FUNCTION_BLOCK SEC_SWITCH_LR_QUARTER_LWORD (* Section-Switcher: Teilbreiten von links und von rechts abschalten, bis 32 Sections, Maske als LWORD im Condensed Work State (2 Bit je Section) *)
  (* Standard: 61499-2; Description: Copyright (c) 2026 Meisterschulen am Ostbahnhof This program and the accompanying materials are made available under the terms of the Eclipse Public License 2.0 which is available at https://www.eclipse.org/legal/epl-2.0/ SPDX-License-Identifier: EPL-2.0 *)
  (* Version 1.1, 2026-11-01, Franz Höpfinger, Meisterschulen am Ostbahnhof, Alle aus und eigener Zaehler 0: LEFT/RIGHT_OFF_DEC uebernimmt zuerst alle abgeschalteten Sections (nach ALL_OFF schaltet Links_Ein von rechts, Rechts_Ein von links zu) *)
  (* Version 1.0, 2026-10-31, Franz Höpfinger, Meisterschulen am Ostbahnhof, initial implementation *)
  PACKAGE logiBUS::sections;
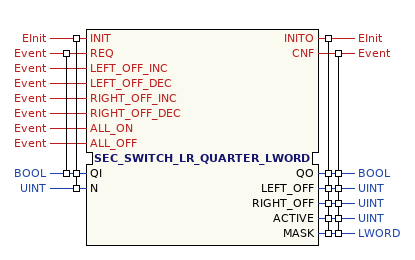
  EVENT_INPUT
    INIT : EInit WITH QI, N; (* Initialisierung, Zaehler auf 0 *)
    REQ WITH QI; (* Maske und Zaehler erneut ausgeben *)
    LEFT_OFF_INC; (* Von links eine Section mehr abschalten *)
    LEFT_OFF_DEC; (* Von links eine Section wieder zuschalten *)
    RIGHT_OFF_INC; (* Von rechts eine Section mehr abschalten *)
    RIGHT_OFF_DEC; (* Von rechts eine Section wieder zuschalten *)
    ALL_ON; (* Alle Sections zuschalten (beide Zaehler 0) *)
    ALL_OFF; (* Alle Sections abschalten (LEFT_OFF = N, RIGHT_OFF = 0) *)
  END_EVENT
  EVENT_OUTPUT
    INITO : EInit WITH QO, LEFT_OFF, RIGHT_OFF, ACTIVE, MASK; (* Initialisierung bestaetigt *)
    CNF WITH QO, LEFT_OFF, RIGHT_OFF, ACTIVE, MASK; (* Zaehler oder Maske neu berechnet *)
  END_EVENT
  VAR_INPUT
    QI : BOOL := TRUE; (* Nur an INIT und REQ: INIT+ aktiv, INIT- deaktiviert (Maske alle frei), REQ- ohne Wirkung *)
    N : UINT; (* Anzahl Sections (1..32, groesser wird auf 32 begrenzt) *)
  END_VAR
  VAR_OUTPUT
    QO : BOOL; (* TRUE = aktiv und Ereignis ausgefuehrt *)
    LEFT_OFF : UINT; (* Anzahl von links abgeschalteter Sections *)
    RIGHT_OFF : UINT; (* Anzahl von rechts abgeschalteter Sections *)
    ACTIVE : UINT; (* Anzahl freier Sections *)
    MASK : LWORD; (* Maske, 2 Bit je Section: 01 frei, 00 gesperrt, 11 nicht vorhanden (Section > N); Bits 1..0 = Section 1 (links) *)
  END_VAR
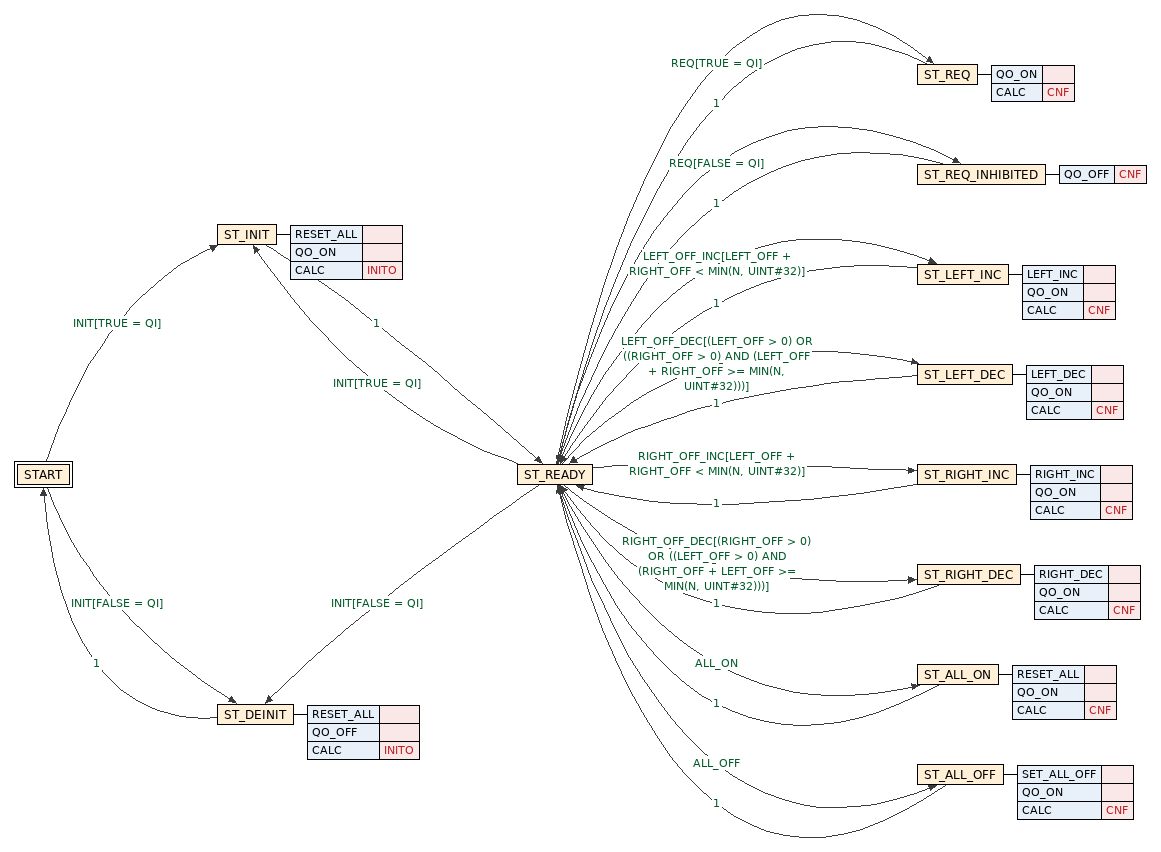
  EC_STATES
    START; (* Nicht initialisiert bzw. deaktiviert *)
    ST_INIT : RESET_ALL, QO_ON, CALC -> INITO; (* INIT+: N uebernehmen, Zaehler 0 *)
    ST_READY; (* Aktiv *)
    ST_DEINIT : RESET_ALL, QO_OFF, CALC -> INITO; (* INIT-: deaktiviert, Maske alle frei *)
    ST_REQ : QO_ON, CALC -> CNF; (* REQ+: Maske und Zaehler ausgeben *)
    ST_REQ_INHIBITED : QO_OFF -> CNF; (* REQ-: nichts aendern, nur melden *)
    ST_LEFT_INC : LEFT_INC, QO_ON, CALC -> CNF;
    ST_LEFT_DEC : LEFT_DEC, QO_ON, CALC -> CNF;
    ST_RIGHT_INC : RIGHT_INC, QO_ON, CALC -> CNF;
    ST_RIGHT_DEC : RIGHT_DEC, QO_ON, CALC -> CNF;
    ST_ALL_ON : RESET_ALL, QO_ON, CALC -> CNF;
    ST_ALL_OFF : SET_ALL_OFF, QO_ON, CALC -> CNF;
  END_STATES
  EC_TRANSITIONS
    START TO ST_INIT := INIT[TRUE = QI];
    START TO ST_DEINIT := INIT[FALSE = QI];
    ST_INIT TO ST_READY := 1;
    ST_DEINIT TO START := 1;
    ST_READY TO ST_INIT := INIT[TRUE = QI];
    ST_READY TO ST_DEINIT := INIT[FALSE = QI];
    ST_READY TO ST_REQ := REQ[TRUE = QI];
    ST_REQ TO ST_READY := 1;
    ST_READY TO ST_REQ_INHIBITED := REQ[FALSE = QI];
    ST_REQ_INHIBITED TO ST_READY := 1;
    ST_READY TO ST_LEFT_INC := LEFT_OFF_INC[LEFT_OFF + RIGHT_OFF < MIN(N, UINT#32)];
    ST_LEFT_INC TO ST_READY := 1;
    ST_READY TO ST_LEFT_DEC := LEFT_OFF_DEC[(LEFT_OFF > 0) OR ((RIGHT_OFF > 0) AND (LEFT_OFF + RIGHT_OFF >= MIN(N, UINT#32)))];
    ST_LEFT_DEC TO ST_READY := 1;
    ST_READY TO ST_RIGHT_INC := RIGHT_OFF_INC[LEFT_OFF + RIGHT_OFF < MIN(N, UINT#32)];
    ST_RIGHT_INC TO ST_READY := 1;
    ST_READY TO ST_RIGHT_DEC := RIGHT_OFF_DEC[(RIGHT_OFF > 0) OR ((LEFT_OFF > 0) AND (RIGHT_OFF + LEFT_OFF >= MIN(N, UINT#32)))];
    ST_RIGHT_DEC TO ST_READY := 1;
    ST_READY TO ST_ALL_ON := ALL_ON;
    ST_ALL_ON TO ST_READY := 1;
    ST_READY TO ST_ALL_OFF := ALL_OFF;
    ST_ALL_OFF TO ST_READY := 1;
  END_TRANSITIONS
  ALGORITHM RESET_ALL IN ST:
LEFT_OFF := 0;
RIGHT_OFF := 0;
  END_ALGORITHM
  ALGORITHM LEFT_INC IN ST:
LEFT_OFF := LEFT_OFF + 1;
  END_ALGORITHM
  ALGORITHM LEFT_DEC IN ST:
(* Alle aus und eigener Zaehler 0: diese Seite uebernimmt zuerst alle
   abgeschalteten Sections, damit beide Seiten nach ALL_OFF zuschalten *)
IF (LEFT_OFF = 0) AND (RIGHT_OFF > 0) AND (LEFT_OFF + RIGHT_OFF >= MIN(N, UINT#32)) THEN
	LEFT_OFF := RIGHT_OFF;
	RIGHT_OFF := 0;
END_IF;
(* Schutz gegen UINT-Unterlauf, zusaetzlich zur ECC-Bedingung *)
IF LEFT_OFF > 0 THEN
	LEFT_OFF := LEFT_OFF - 1;
END_IF;
  END_ALGORITHM
  ALGORITHM RIGHT_INC IN ST:
RIGHT_OFF := RIGHT_OFF + 1;
  END_ALGORITHM
  ALGORITHM RIGHT_DEC IN ST:
(* Alle aus und eigener Zaehler 0: diese Seite uebernimmt zuerst alle
   abgeschalteten Sections, damit beide Seiten nach ALL_OFF zuschalten *)
IF (RIGHT_OFF = 0) AND (LEFT_OFF > 0) AND (RIGHT_OFF + LEFT_OFF >= MIN(N, UINT#32)) THEN
	RIGHT_OFF := LEFT_OFF;
	LEFT_OFF := 0;
END_IF;
(* Schutz gegen UINT-Unterlauf, zusaetzlich zur ECC-Bedingung *)
IF RIGHT_OFF > 0 THEN
	RIGHT_OFF := RIGHT_OFF - 1;
END_IF;
  END_ALGORITHM
  ALGORITHM SET_ALL_OFF IN ST:
LEFT_OFF := MIN(N, UINT#32);
RIGHT_OFF := 0;
  END_ALGORITHM
  ALGORITHM QO_ON IN ST:
QO := TRUE;
  END_ALGORITHM
  ALGORITHM QO_OFF IN ST:
QO := FALSE;
  END_ALGORITHM
  ALGORITHM CALC IN ST:
VAR_TEMP
	nEff : UINT; // N begrenzt auf 32
	lastOn : UINT; // letzte freie Section
	freeAll : LWORD; // ACTIVE Paare Einsen
	notThere : LWORD; // 11 fuer Sections > N
END_VAR
(* 1. Begrenzung auf gueltigen Bereich 0..32 *)
nEff := MIN(N, UINT#32);
LEFT_OFF := MIN(LEFT_OFF, nEff);
RIGHT_OFF := MIN(RIGHT_OFF, nEff - LEFT_OFF);
(* 2. Aktive Sections berechnen *)
lastOn := nEff - RIGHT_OFF;
ACTIVE := lastOn - LEFT_OFF;
(* 3. Maske ohne Schleife: freie Sections 01 (ACTIVE Paare ab LEFT_OFF, nur unteres Bit),
   Sections ueber N 11, alle anderen 00 *)
IF ACTIVE >= UINT#32 THEN
	freeAll := LWORD#16#FFFFFFFFFFFFFFFF;
ELSE
	freeAll := NOT SHL(LWORD#16#FFFFFFFFFFFFFFFF, 2 * ACTIVE);
END_IF;
IF nEff >= UINT#32 THEN
	notThere := LWORD#0;
ELSE
	notThere := SHL(LWORD#16#FFFFFFFFFFFFFFFF, 2 * nEff);
END_IF;
MASK := (SHL(freeAll, 2 * LEFT_OFF) AND LWORD#16#5555555555555555) OR notThere;
  END_ALGORITHM
  SERVICE APPLICATION/SWITCHER (* QI wirkt nur an INIT und REQ (INIT+/INIT-, REQ+/REQ-). Tasten, ALL_ON und ALL_OFF wirken im aktiven Zustand ohne QI. *)
    SEQUENCE normal_initialization (* INIT mit QI = TRUE: N uebernehmen, alle Sections frei *)
      APPLICATION.INIT+(N) -> APPLICATION.INITO+(LEFT_OFF,RIGHT_OFF,ACTIVE,MASK);
    END_SEQUENCE
    SEQUENCE re_initialization (* INIT+ im aktiven Zustand: neu initialisieren, Zaehler 0 *)
      APPLICATION.INIT+(N) -> APPLICATION.INITO+(LEFT_OFF,RIGHT_OFF,ACTIVE,MASK);
    END_SEQUENCE
    SEQUENCE termination (* INIT mit QI = FALSE: deaktiviert, Maske alle frei *)
      APPLICATION.INIT-() -> APPLICATION.INITO-(LEFT_OFF,RIGHT_OFF,ACTIVE,MASK);
    END_SEQUENCE
    SEQUENCE termination_without_initialization (* INIT- auch vor INIT+ wird mit INITO- beantwortet (INIT-Kette haengt nicht) *)
      APPLICATION.INIT-() -> APPLICATION.INITO-(LEFT_OFF,RIGHT_OFF,ACTIVE,MASK);
    END_SEQUENCE
    SEQUENCE request (* Maske und Zaehler erneut ausgeben *)
      APPLICATION.REQ+() -> APPLICATION.CNF+(LEFT_OFF,RIGHT_OFF,ACTIVE,MASK);
    END_SEQUENCE
    SEQUENCE request_inhibited (* REQ mit QI = FALSE: nichts aendern *)
      APPLICATION.REQ-() -> APPLICATION.CNF-();
    END_SEQUENCE
    SEQUENCE left_off_increment (* Von links eine Section mehr abschalten *)
      APPLICATION.LEFT_OFF_INC() -> APPLICATION.CNF+(LEFT_OFF,RIGHT_OFF,ACTIVE,MASK);
    END_SEQUENCE
    SEQUENCE left_off_increment_at_limit (* Alle Sections schon aus: keine Reaktion *)
      APPLICATION.LEFT_OFF_INC();
    END_SEQUENCE
    SEQUENCE left_off_decrement (* Von links eine Section wieder zuschalten *)
      APPLICATION.LEFT_OFF_DEC() -> APPLICATION.CNF+(LEFT_OFF,RIGHT_OFF,ACTIVE,MASK);
    END_SEQUENCE
    SEQUENCE left_off_decrement_at_zero (* LEFT_OFF = 0: keine Reaktion *)
      APPLICATION.LEFT_OFF_DEC();
    END_SEQUENCE
    SEQUENCE right_off_increment (* Von rechts eine Section mehr abschalten *)
      APPLICATION.RIGHT_OFF_INC() -> APPLICATION.CNF+(LEFT_OFF,RIGHT_OFF,ACTIVE,MASK);
    END_SEQUENCE
    SEQUENCE right_off_decrement (* Von rechts eine Section wieder zuschalten *)
      APPLICATION.RIGHT_OFF_DEC() -> APPLICATION.CNF+(LEFT_OFF,RIGHT_OFF,ACTIVE,MASK);
    END_SEQUENCE
    SEQUENCE all_on (* Alle Sections zuschalten *)
      APPLICATION.ALL_ON() -> APPLICATION.CNF+(LEFT_OFF,RIGHT_OFF,ACTIVE,MASK);
    END_SEQUENCE
    SEQUENCE all_off (* Alle Sections abschalten (LEFT_OFF = N) *)
      APPLICATION.ALL_OFF() -> APPLICATION.CNF+(LEFT_OFF,RIGHT_OFF,ACTIVE,MASK);
    END_SEQUENCE
    SEQUENCE event_before_initialization (* REQ, Tasten, ALL_ON/ALL_OFF vor INIT+ bzw. nach INIT-: keine Reaktion *)
      APPLICATION.REQ();
    END_SEQUENCE
    SEQUENCE left_on_after_all_off (* Nach ALL_OFF: LEFT_OFF_DEC schaltet die rechte Section N zu, dann N-1 ... *)
      APPLICATION.LEFT_OFF_DEC() -> APPLICATION.CNF+(LEFT_OFF,RIGHT_OFF,ACTIVE,MASK);
    END_SEQUENCE
    SEQUENCE right_on_after_all_off (* Nach ALL_OFF: RIGHT_OFF_DEC schaltet die linke Section 1 zu, dann 2 ... *)
      APPLICATION.RIGHT_OFF_DEC() -> APPLICATION.CNF+(LEFT_OFF,RIGHT_OFF,ACTIVE,MASK);
    END_SEQUENCE
  END_SERVICE
END_FUNCTION_BLOCK
